Staubli VAL3: dioItem.pjx

--- dioItem.pjx ---
Parameters version=s8.10.3Cs9_BS2093 stackSize=5000 millimeterUnit=true
Program file=start.pgx
Program file=stop.pgx
Data file=dioItem.dtx

--- dioItem.dtx ---
public string sComment
public dio dDio

--- start.pgx ---
program start()
begin
end

--- stop.pgx ---
program stop()
begin
end
